(* IEC 61131-3 sources: Lasal-MCP/examples/SampleSource/4_PumpControlSchemeSolution/Stations/Terminal/HMI/Class/_SyncTimeHMI, 1 file *)

(* ---- _SyncTimeHMI.st ---- *)
(*!
<Class
	Name               = "_SyncTimeHMI"
	Revision           = "1.1"
	RealtimeTask       = "false"
	CyclicTask         = "false"
	BackgroundTask     = "false"
	Sigmatek           = "true"
	OSInterface        = "false"
	HighPriority       = "false"
	Automatic          = "false"
	UpdateMode         = "Prescan"
	SharedCommandTable = "true"
	Objectsize         = "(540,180)"
	Comment            = "class reads date and time from two clients (within the adjusted zycletime)&#13;&#10;and writes these values to the servers">
	<Channels>
		<Server Name="sSyncDate" Visualized="true" Initialize="false" WriteProtected="true" Retentive="false" Comment="server for sync date"/>
		<Server Name="sSyncTime" Visualized="true" Initialize="false" WriteProtected="true" Retentive="false" Comment="server for sync time"/>
		<Client Name="ActDate" Required="true" Internal="false" Comment="actual date"/>
		<Client Name="ActTime" Required="true" Internal="false" Comment="actual time"/>
	</Channels>
	<Dependencies>
		<Files>
			<File Path=".\Class\_SyncTimeHMI\_SyncTimeHMI_de.pdf"/>
			<File Path=".\Class\_SyncTimeHMI\_SyncTimeHMI_en.pdf"/>
		</Files>
	</Dependencies>
	<RevDoku>
		<Owner Company="Sigmatek"/>
		<Dokumentation Revision="1.1" Date="2016-10-10" Author="HubChr" Company="Sigmatek" Description="Added documentation pdfs."/>
		<Dokumentation Revision="1.0" Date="2015-11-11" Author="hötant" Company="Sigmatek" Description="creation of class"/>
	</RevDoku>
</Class>
*)
_SyncTimeHMI : CLASS
  //Servers:
	sSyncDate 	: SvrChCmd_HDINT;
	sSyncTime 	: SvrCh_HDINT;
  //Clients:
	ActDate 	: CltCh_HDINT;
	ActTime 	: CltCh_HDINT;
  //Variables:
  //Functions:

	FUNCTION VIRTUAL GLOBAL sSyncDate::Read
		VAR_OUTPUT
			output (EAX) 	: HDINT;
		END_VAR;

	FUNCTION VIRTUAL GLOBAL sSyncTime::Read
		VAR_OUTPUT
			output (EAX) 	: HDINT;
		END_VAR;
  //Tables:
	FUNCTION @STD
		VAR_OUTPUT
			ret_code	: CONFSTATES;
		END_VAR;
	FUNCTION GLOBAL TAB @CT_;
END_CLASS;

FUNCTION VIRTUAL GLOBAL _SyncTimeHMI::sSyncDate::Read
	VAR_OUTPUT
		output (EAX) 	: HDINT;
	END_VAR

	output := sSyncDate := ActDate := ActDate.Read();

END_FUNCTION

FUNCTION VIRTUAL GLOBAL _SyncTimeHMI::sSyncTime::Read
	VAR_OUTPUT
		output (EAX) 	: HDINT;
	END_VAR

	output := sSyncTime :=ActTime :=  ActTime.Read();

END_FUNCTION
